// TIA Portal project "PLC_hackathon_2026_V21" (V21)

(* hardware
DEVICE "S71500/ET200MP station_1"  S7-1500 station
   slot 0: "Rail_0"  Rack  6ES7 590-1***0-0AA0
   slot 1: "PLC_1"  CPU 1515-2 PN  6ES7 515-2AM01-0AB0  V2.6
      slot 3: "CPU display_1"  6ES7591-1BA00-0AA0
DEVICE "PC-System_1"  SIMATIC PC station
   slot 0: "SIMATIC PC station"  Rail  SIMATIC PC-Station  V1.0
      slot 125: "Stationmanager"  Station_Manager  V6.0.4
   slot 1: "HMI_RT_1"  WinCC RT Advanced  6AV2 104-0xxxx-xxxx  17.0.0.0
      slot 33792: "Host interface"  Host interface
   slot 2: "IE general_1"  IE General  IE_CP  V8.2.0
*)

// ===== PLC "PLC_1"  CPU 1515-2 PN =====
// protected blocks, not shown: "Crane_manipulation"

VAR_GLOBAL   // PLC tag table "Default tag table"
   "x_position" AT %MB104 : SInt;
   "y_position" AT %MB105 : SInt;
   "bay_ID" AT %MB106 : USInt;
   "number_of_manipulations" AT %MD107 : UDInt;
   "time" AT %MD112 : Real;
END_VAR

VAR_GLOBAL   // PLC tag table "Crane_command"
   "new_x_position" AT %MB100 : SInt;   // X position for the move command
   "new_y_position" AT %MB101 : SInt;   // Y position for the move command
   "new_bay_ID" AT %MB102 : USInt;   // Bay ID for the move command
   "new_command_ID" AT %MB103 : USInt;   // ID of the command
END_VAR

TYPE "typeCmd"
   STRUCT
      Cmd : USInt;   // 0 none, 1 lift, 2 put down, 3 move to (X,Y,Bay), 10 reset
      X : SInt;   // 0..3 (for lift/put: current crane x)
      Y : SInt;   // 0..11 (for lift/put: current crane y)
      Bay : USInt;   // 0 ship, 1 yard
      Src : USInt;   // origin: 1 AUTO, 2 SEMI, 3 MANUAL, 4 INIT(reset)
      TrIdx : Int;   // plan transfer index (0 = not from plan)
      Phase : USInt;   // 0 move-to-src, 1 lift, 2 move-to-dst, 3 put (only if TrIdx>0)
   END_STRUCT;
END_TYPE

TYPE "typeTransfer"
   STRUCT
      Kind : USInt;   // 1 unload (Bay0->Bay1), 2 load (Bay1->Bay0)
      Id : UInt;   // container ID
      ListIdx : Int;   // index into UList (Kind 1) or LList (Kind 2)
      SrcX : SInt;
      SrcY : SInt;
      SrcBay : USInt;
      DstX : SInt;
      DstY : SInt;
      DstBay : USInt;
      CumT_ds : DInt;   // predicted total time after this transfer, deciseconds, incl. BaseT_ds
      CumM : DInt;   // predicted total manipulations after this transfer, incl. BaseM
   END_STRUCT;
END_TYPE

DATA_BLOCK "Current_state_of_Bay0"   // DB10
{ S7_Optimized_Access := 'TRUE' }
VERSION : 0.1
   VAR
      Bay0 : Array[0..3, 0..11] of UInt;
   END_VAR
BEGIN
   Bay0[0,0] := 123;
   Bay0[0,1] := 326;
   Bay0[0,2] := 987;
END_DATA_BLOCK

DATA_BLOCK "Current_state_of_Bay1"   // DB11
{ S7_Optimized_Access := 'TRUE' }
VERSION : 0.1
   VAR
      Bay1 : Array[0..3, 0..11] of UInt;
   END_VAR
BEGIN
   Bay1[0,1] := 246;
   Bay1[0,7] := 675;
   Bay1[1,5] := 777;
END_DATA_BLOCK

DATA_BLOCK "From_Bay0_to_Bay1"   // DB20
{ S7_Optimized_Access := 'TRUE' }
VERSION : 0.1
   VAR
      IDs_of_the_containers : Array[1..48] of UInt;
   END_VAR
BEGIN
   IDs_of_the_containers[12] := 0;
   IDs_of_the_containers[18] := 0;
   IDs_of_the_containers[4] := 444;
   IDs_of_the_containers[1] := 111;
   IDs_of_the_containers[2] := 222;
   IDs_of_the_containers[3] := 333;
   IDs_of_the_containers[5] := 555;
   IDs_of_the_containers[6] := 666;
   IDs_of_the_containers[7] := 777;
END_DATA_BLOCK

DATA_BLOCK "From_Bay1_to_Bay0"   // DB21
{ S7_Optimized_Access := 'TRUE' }
VERSION : 0.1
   VAR
      Bay1_IDs_of_the_containers : Array[1..48] of UInt;
   END_VAR
BEGIN
   Bay1_IDs_of_the_containers[15] := 0;
   Bay1_IDs_of_the_containers[22] := 0;
   Bay1_IDs_of_the_containers[1] := 123;
   Bay1_IDs_of_the_containers[2] := 124;
   Bay1_IDs_of_the_containers[3] := 125;
END_DATA_BLOCK

DATA_BLOCK "World"   // DB100
{ S7_Optimized_Access := 'TRUE' }
VERSION : 0.1
   VAR
      Bay0 : Array[0..3, 0..11] of UInt;   // working copy of the ship (FB10 INIT copy / OB30 lift-put effect)
      Bay1 : Array[0..3, 0..11] of UInt;   // working copy of the yard
      CraneX : SInt;   // crane x after last completed command
      CraneY : SInt;
      CraneBay : USInt := 1;
      Carried : UInt;   // ID on the hook (0 = none)
      Busy : Bool;   // command issued to FB1, not finished yet
      BusyTicks : Int;   // OB30 ticks since issue (watchdog)
      ActCmd : "typeCmd";   // command currently executing
      NextCmd : "typeCmd";   // staged command (valid when CmdReady)
      CmdReady : Bool;   // handshake: FB10 sets (last) / OB30 clears
      Permit : Bool;   // OB30 may issue NextCmd
      DoneSeq : UDInt;   // +1 per completed command
      LastDone : "typeCmd";   // last completed command
      Fault : Word;   // OB30-detected alarms (bit = alarm bit)
      FaultCmd : "typeCmd";   // command rejected by CheckCmd
      UList : Array[1..48] of UInt;   // copy of DB20 (unload list)
      UState : Array[1..48] of USInt;   // 0 pending, 1 done, 2 skipped
      LList : Array[1..48] of UInt;   // copy of DB21 (load list)
      LState : Array[1..48] of USInt;   // as UState
      N : Int;   // non-zero entries in DB20 + DB21 (for J)
      Plan : Array[1..96] of "typeTransfer";   // written by the planner
      PlanLen : Int;
      PlanValid : Bool;
      PlanVariant : Int;
      PredT_ds : DInt;
      PredM : DInt;
      PredJ : Real;
      BaseT_ds : DInt;   // ROUND(T*10) at plan request
      BaseM : DInt;   // M at plan request
      PlanIdx : Int := 1;   // done pointer: transfer being executed
      Phase : USInt;   // done pointer: next phase of PlanIdx to complete
      StageIdx : Int := 1;   // staging cursor (transfer)
      StagePhase : USInt;   // staging cursor (phase)
      BalL : Int;   // ship count x in {0,1}
      BalR : Int;   // ship count x in {2,3}
      BalF : Int;   // ship count y in 0..5
      BalA : Int;   // ship count y in 6..11
      CfgOrderMode : USInt := 1;   // 0 free, 1 per-list order, 2 strict (set by FB10 from HMI_IF before each plan)
      CfgBalLimit : Int := 5;
      CfgBalMode : USInt;   // 0 x-halves only, 1 also y-halves
      CfgMMode : USInt := 0;   // manipulation count model (CONTRACT 4.1); v1.7: 0 = spec rule (diagonal = 2), 2 = FB1 (+1 per move command)
      CfgVariants : Int := 4;
      CfgAlpha : Array[1..4] of Int;   // v1.7: retuned for CfgMMode 0 (v1.3 mode 2: [0, 100, 200, 300])
      CfgStepsPerCall : Int := 1;
      CfgTimeoutTicks : Int := 10;   // FB1 watchdog in OB30 ticks (1 s)
      OB30Ticks : UDInt;
      MSpec : UDInt;   // manipulations by the spec rule (OB30): +1 per changed axis, +1 lift/put ---- v1.3: improve phase (CONTRACT 4.8) and lower bound (4.9) ----
      CfgImproveEvals : DInt := 3000;   // local-search evaluations after the greedy (0 = off)
      CfgImproveDist : Int := 0;   // max |i-j| of a move (0 = unlimited)
      CfgImprovePerCall : Int := 1;   // evaluations per OB1 call (per-call work bound)
      PredJ0 : Real;   // J of the greedy winner before the improve phase
      LbT_ds : DInt;   // lower bound of the final T (incl. BaseT_ds), deciseconds
      LbM : DInt;   // lower bound of the final M (incl. BaseM)
      LbJ : Real;   // lower bound of J (no plan can be better)
      ImpEvals : DInt;   // improve phase: evaluations done (last plan)
      ImpAccepts : DInt;   // improve phase: accepted improvements (last plan) ---- v1.4: exact order feasibility (CONTRACT 4.10) and SLOT phase (4.11) ----
      CfgSlotSweeps : Int := 10;   // drop-cell local search sweeps after IMPROVE (0 = off)
      SlotAccepts : DInt;   // SLOT phase: accepted drop-cell changes (last plan)
      OrderFeasible : Bool;   // last plan job: the requested order mode is feasible (exact DP) ---- v1.5 (judge round 2 R2-J1): relaxed balance rule on a ship that starts out of balance ----
      BalCeil : Int;   // 0 = step rule; > CfgBalLimit: while |L-R| > CfgBalLimit a step may go up to BalCeil ---- v1.6 (judge round 3 R3-E3): relaxed ceiling search ----
      CfgRelaxMin : Bool;   // FALSE: relaxed fallback uses BalCeil = start imbalance at once; TRUE: ascending CfgBalLimit+1 .. start imbalance (smallest feasible, costs J)
   END_VAR
BEGIN
   CfgAlpha[1] := 0;
   CfgAlpha[2] := 75;
   CfgAlpha[3] := 125;
   CfgAlpha[4] := 200;
END_DATA_BLOCK

DATA_BLOCK "HMI_IF"   // DB101
{ S7_Optimized_Access := 'TRUE' }
VERSION : 0.1
// ---- Buttons / inputs (HMI writes; FB10 resets button bits after evaluating them) ----
   VAR
      SwOn : Bool;   // main switch level (HMI InvertBit), TRUE = ON
      BtnInit : Bool;   // INITIAL STATE (POCETNO STANJE)
      BtnAuto : Bool;
      BtnSemi : Bool;
      BtnManual : Bool;
      BtnStart : Bool;
      BtnStop : Bool;
      BtnAck : Bool;
      BtnStep : Bool;   // SEMI: run the next manipulation
      BtnManExec : Bool;   // MANUAL: execute ManCmd
      ManCmd : USInt;   // 1 lift, 2 put down, 3 move, 10 reset
      ManX : SInt;   // 0..3
      ManY : SInt;   // 0..11
      ManBay : USInt;   // 0 ship, 1 yard
      CfgOrderMode : USInt := 1;   // 0 free, 1 per-list order (default, hedge), 2 strict; FB10 falls back 2->1->0 if infeasible
      CfgSemiPerTransfer : Bool;   // SEMI click = one command (FALSE) or one transfer (TRUE)
      CfgBalMode : USInt;   // 0 x-halves, 1 also y-halves
      AlarmHmiAck : Word;   // WinCC 'Acknowledgement tag': alarm acknowledged in the alarm view (= POTVRDA); FB10 resets it ---- Indicators (FB10 writes every OB1 cycle) ----
      State : USInt;   // 0 OFF,1 INIT,2 READY,3 RUNNING,4 PAUSED,5 ALARM,6 DONE,7 PLANNING
      Mode : USInt := 1;   // 1 AUTO, 2 SEMI, 3 MANUAL
      LampOn : Bool;
      LampOff : Bool;
      LampReady : Bool;
      LampAuto : Bool;
      LampSemi : Bool;
      LampManual : Bool;
      LampRunning : Bool;
      LampAlarm : Bool;
      LampDone : Bool;
      Initialized : Bool;
      CraneBusy : Bool;
      Planning : Bool;
      StepWaiting : Bool;   // SEMI is waiting for a click
      "M" : UDInt;   // v1.7: M by the spec rule (x and y change = 2) = World.MSpec (primary)
      T : Real;   // = "time" (MD112) working time [s]
      J : Real;   // v1.7: 0.5*T/(76*N) + 0.5*M/(4*N) with the spec M (primary)
      MSpec : UDInt;   // = M (spec rule, computed in OB30); kept for compatibility
      JSpec : Real;   // = J (spec rule); kept for compatibility
      MFb1 : UDInt;   // v1.7: FB1's own counter "number_of_manipulations" (MD107, +1 per command)
      JFb1 : Real;   // v1.7: J with MFb1 (secondary)
      OrderModeAct : USInt;   // order mode actually used by the last plan (after fallback)
      OrderFallback : Bool;   // v1.4: preferred order/balance mode infeasible, plan uses a weaker one
      SlotAccepts : DInt;   // v1.4: SLOT phase accepted drop-cell changes (last plan)
      N : Int;
      PredM : DInt;
      PredT : Real;
      PredJ : Real;
      PredJ0 : Real;   // v1.3: greedy J before the improve phase
      LbJ : Real;   // v1.3: lower bound of J (no plan can be better)
      GapPct : Real;   // v1.3: (PredJ / LbJ - 1) * 100
      ImpGainPct : Real;   // v1.3: (1 - PredJ / PredJ0) * 100 = gain of the improve phase
      ImpEvals : DInt;   // v1.3: improve-phase evaluations of the last plan
      PlanProgress : Int;   // v1.3: planner progress 0..100 % (improve phase)
      PlanVariant : Int;
      TrDone : Int;
      TrTotal : Int;
      UDone : Int;
      UTotal : Int;
      LDone : Int;
      LTotal : Int;
      CraneX : SInt;
      CraneY : SInt;
      CraneBay : USInt;
      CraneGX : Int;   // global column: x+6 if bay 0 else x (0..9)
      Carried : UInt;
      CurCmd : USInt;
      CurX : SInt;
      CurY : SInt;
      CurBay : USInt;
      CurId : UInt;
      CurKind : USInt;   // 1 unload, 2 load, 0 none
      CurPhase : USInt;
      Cell0 : Array[0..47] of UInt;   // Bay0 IDs, index x*12+y
      Cell1 : Array[0..47] of UInt;   // Bay1 IDs, index x*12+y
      CellSt0 : Array[0..47] of USInt;   // colour code 0..7
      CellSt1 : Array[0..47] of USInt;
      UList : Array[1..48] of UInt;
      LList : Array[1..48] of UInt;
      UState : Array[1..48] of USInt;   // 0 pending, 1 done, 2 skipped, 3 in progress
      LState : Array[1..48] of USInt;
      BalL : Int;
      BalR : Int;
      BalDiff : Int;   // BalL - BalR
      BalF : Int;
      BalA : Int;
      BalOk : Bool;   // |BalDiff| <= 5
      AlarmWord : Word;   // alarm bits (CONTRACT 3.3)
      AlarmAckWord : Word;   // WinCC 'PLC acknowledgement tag' = NOT AlarmWord (one ACK clears PLC and HMI)
      AlarmId : UInt;
      AlarmWord2 : Word;   // v1.4: extra alarm bits: bit 0 = list order abandoned (warning); v1.5 bit 1 = relaxed balance rule (ship loaded unbalanced)
      AlarmUId : UInt;   // v1.4: first unload-list ID that is not in Bay 0 (alarm bit 3)
      AlarmUCnt : Int;   // number of such IDs
      AlarmLId : UInt;   // v1.4: first load-list ID that is not in Bay 1 (alarm bit 4)
      AlarmLCnt : Int;
      AlarmX : SInt;
      AlarmY : SInt;
      AlarmBay : USInt;
      AlarmHist : Array[0..15] of Int;   // alarm bit numbers of the last 16 raises, [0] newest
      AlarmHistSeq : UDInt;
      OB30Ticks : UDInt;
      Heartbeat : Bool;   // toggles each OB30 tick
   END_VAR
BEGIN
END_DATA_BLOCK

DATA_BLOCK "Crane_Control_DB"   // DB110
{ S7_Optimized_Access := 'TRUE' }
VERSION : 0.1
// stored: InstanceOfName Crane_Control
"Crane_Control"
BEGIN
END_DATA_BLOCK

// folder: Constants

DATA_BLOCK "Global_constants"   // DB1
{ S7_Optimized_Access := 'TRUE' }
VERSION : 0.1
   VAR
      container_width_in_m : Real := 2.3;   // Container width in meters
      container_length_in_m : Real := 6.0;   // Container length in meters
      velocity_of_the_crane_in_m_per_s : Real := 1.0;   // Velocity of the crane in meters per second
      time_to_lift_a_container_in_s : Real := 20.0;   // Time needed to lower the hook, hook up a container and lift it in seconds
      time_to_put_down_a_container_in_s : Real := 20.0;   // Time needed to put down a container, release it, and lift up the hook in seconds
   END_VAR
BEGIN
END_DATA_BLOCK

// folder: (top level)

FUNCTION_BLOCK "Crane_Control"   // FB10, SCL
TITLE = Container crane control (FB10, called from OB1)
{ S7_Optimized_Access := 'TRUE' }
VERSION : 0.1
// FB10 decides WHAT the crane does; OB30 decides WHEN (CONTRACT 3.4).
//   - HMI buttons, modes AUTO / SEMI-AUTO / MANUAL
//   - state machine OFF / INIT / READY / RUNNING / PAUSED / ALARM / DONE / PLANNING
//   - INIT: reset FB1, copy DB10/DB11, validate lists and IDs, call the planner
//   - stages plan commands into "World".NextCmd (handshake CmdReady / Permit)
//   - tracks progress (done pointer), list states, ship balance, alarms
//   - writes every indicator of "HMI_IF"
//   FB10 never calls FB1 and never writes MB100..MB103; FB1 tags are read-only here.
   VAR
      Planner : "Crane_Planner";   // planning algorithm (FB11, CONTRACT 4)
      PlanReq : Bool;   // Req input of the planner
      PlanFinished : Bool;   // planner job ended, result not yet consumed
      PlanOk : Bool;
      PlanErr : Int;
      PlanStep : Int;   // PLANNING sub-step
      PlanCrX : SInt;   // crane position at plan request
      PlanCrY : SInt;
      PlanCrBay : USInt;
      FirstPh : Array[1..96] of USInt;   // first phase of each transfer (1 = move-to-src skipped)
      State : USInt;   // 0 OFF,1 INIT,2 READY,3 RUNNING,4 PAUSED,5 ALARM,6 DONE,7 PLANNING
      PrevState : USInt;   // state to return to after ALARM + ACK
      OffState : USInt;   // state before OFF
      Mode : USInt := 1;   // 1 AUTO, 2 SEMI, 3 MANUAL
      PendMode : USInt;   // mode press waiting to be applied
      Initialized : Bool;
      InitStep : Int;   // INIT sub-step
      InitSeq : UDInt;   // DoneSeq when the INIT reset was staged
      SeenSeq : UDInt;   // last "World".DoneSeq processed
      Resync : Bool;   // re-align staging cursor to done pointer before staging
      SemiTokens : Int;   // SEMI: commands still allowed by BtnStep
      AlarmLatch : Word;   // latched alarm bits (CONTRACT 3.3)
      AlarmPrev : Word;   // for raise-edge detection (history)
      AlarmHistM : Array[0..15] of UDInt;   // M at each history entry (parallel to HMI_IF.AlarmHist)
      AlarmHistT : Array[0..15] of Real;   // T [s] at each history entry
      FirstScan : Bool := TRUE;
      Snap0 : Array[0..3, 0..11] of UInt;   // DB10 as last seen: external online edits are adopted into World
      Snap1 : Array[0..3, 0..11] of UInt;   // DB11 as last seen
      PendStep : Bool;   // SEMI: latched NEXT STEP click (kept while FB1 is busy)
      ReplanAfterPut : Bool;   // destination re-targeted after ACK: replan after that put
      CfgOrdHmi : USInt := 1;   // CfgOrderMode last taken from the HMI (preferred mode)
      CfgBalHmi : USInt;   // CfgBalMode last taken from the HMI
      OrdFallback : Bool;   // next plan request is a fallback retry (keep World.Cfg*) v1.4: DB10/DB11 are kept as the live state; copy of the loaded data for POÄŒETNO STANJE
      InitBay0 : Array[0..3, 0..11] of UInt;
      InitBay1 : Array[0..3, 0..11] of UInt;
      HaveInit : Bool;   // InitBay0/1 valid
      ExtEdit : Bool;   // v1.6: not used any more (NewCnt / ObstCnt), kept for the interface
      NoCellWarn : Bool;   // v1.5: bit 7 raised by the ACK re-target (MANUAL needed): not blocking
      BalD0 : Int;   // v1.5 (R2-J1): |L-R| of the ship as loaded at INIT v1.6 (judge round 3 R3-E1 / R3-J1): obstacle edits during a job are not a new data set
      JobActive : Bool;   // a plan or MANUAL command completed since the last INIT
      EditMark : Array[0..95] of Bool;   // cell (bay*48 + x*12 + y) edited online since the last INIT
      EditNew : Array[0..95] of Bool;   // ... and that edit was made while no job was in progress
      EditVal : Array[0..95] of UInt;   // value of the cell before the edit (written back = unmarked)
      NewCnt : Int;   // marked cells edited with no job in progress (new data)
      ObstCnt : Int;   // marked cells edited during a job (obstacles)
   END_VAR
   VAR_TEMP
      visSt0 : Array[0..47] of USInt;   // display colours built privately
      visSt1 : Array[0..47] of USInt;
      bInit : Bool;   // button snapshots (HMI bits are reset at once)
      bAuto : Bool;
      bSemi : Bool;
      bManual : Bool;
      bStart : Bool;
      bStop : Bool;
      bAck : Bool;
      bStep : Bool;
      bManExec : Bool;
      i : Int;
      j : Int;
      k : Int;
      x : Int;
      y : Int;
      "b" : Int;
      id : UInt;
      found : Bool;
      found0 : Bool;
      found1 : Bool;
      cnt : Int;
      cnt2 : Int;
      pu : Int;
      pl : Int;
      seq : UDInt;
      last : "typeCmd";
      cur : "typeCmd";
      blocking : Bool;
      hadFault : Bool;
      carriedOk : Bool;
      newBits : Word;
      newFault : Word;
      tc : Array[0..95] of UInt;   // INIT: all cells, index bay*48 + x*12 + y
      tl : Array[1..96] of UInt;   // INIT: UList (1..48) then LList (49..96)
      ts : Array[1..96] of USInt;   // INIT: states of tl
      rN : Real;
      curValid : Bool;
      tr : "typeTransfer";
      unbal : Bool;   // ship out of balance now (alarm bit 0 condition)
      semiGo : Bool;   // SEMI NEXT STEP in READY / PAUSED = START + one step
      faultWas : Word;   // World.Fault at ACK
      planPut : Bool;   // completed PUT belongs to the plan
      bestT : Int;   // re-target: best travel time [ds]
      bestX : Int;
      bestY : Int;
      candT : Int;
      nL : Int;
      nR : Int;
      nF : Int;
      nA : Int;
      okBal : Bool;
      dstB : USInt;
      noCell : Bool;   // ACK: rejected plan put could not be re-targeted
      extE : Bool;   // INIT: DB10/DB11 differ from the last mirrored state
      noJob : Bool;   // v1.6: no job in progress (an online edit is new data)
      dbv : UInt;   // v1.6 region 2a: DB10/DB11 cell
      snv : UInt;   // Snap cell
      wv : UInt;   // World cell v1.6 (judge round 3 R3-E2): order feasibility of the ACK re-target (bit-parallel FtMask[0,0])
      ft0 : DWord;   // bit L: the remaining lists stay feasible from L ship containers in x 0..1
      ftNu : Int;   // remaining pending unloads (list order)
      ftNl : Int;   // remaining pending loads (without the one on the hook)
      ftS0 : Int;   // ship count after the put
      ftY0 : Int;   // yard count
      ftCeil : Int;   // ceiling of this try: 0 step rule, > 0 relaxed, -1 skip, -2 no filter
      ftTry : Int;
      ftUse : Bool;   // filter possible (ship put, preferred order 1 / 2)
      ftSide : Array[1..48] of Bool;   // pending unload i (list order) stands in x 0..1
      ftPrev : Array[0..48] of DWord;   // FtMask row i + 1
      ftCur : Array[0..48] of DWord;   // FtMask row i
      ftK : Array[0..4, 0..48] of DWord;   // per ship total: 0 end state, 1 unload left, 2 unload right, 3 load left, 4 load right
      ftTot : Int;
      ftL : Int;
      ftR : Int;
      ftD : Int;
      ftD2 : Int;
      ftM : DWord;
      ftBit : DWord;
      listsNew : Bool;   // v1.6 INIT: DB20/DB21 differ from the lists of the last load
   END_VAR
BEGIN
   REGION 0 First scan after PLC start
       IF #FirstScan THEN
           FOR #i := 0 TO 15 DO
               "HMI_IF".AlarmHist[#i] := -1;      // -1 = empty history entry
           END_FOR;
           #Mode := 1;                            // default AUTO
           #State := 0;
           #FirstScan := FALSE;
       END_IF;
   END_REGION

   REGION 1 HMI buttons: snapshot and reset
       #bInit := "HMI_IF".BtnInit;       "HMI_IF".BtnInit := FALSE;
       #bAuto := "HMI_IF".BtnAuto;       "HMI_IF".BtnAuto := FALSE;
       #bSemi := "HMI_IF".BtnSemi;       "HMI_IF".BtnSemi := FALSE;
       #bManual := "HMI_IF".BtnManual;   "HMI_IF".BtnManual := FALSE;
       #bStart := "HMI_IF".BtnStart;     "HMI_IF".BtnStart := FALSE;
       #bStop := "HMI_IF".BtnStop;       "HMI_IF".BtnStop := FALSE;
       #bAck := "HMI_IF".BtnAck;         "HMI_IF".BtnAck := FALSE;
       #bStep := "HMI_IF".BtnStep;       "HMI_IF".BtnStep := FALSE;
       #bManExec := "HMI_IF".BtnManExec; "HMI_IF".BtnManExec := FALSE;
       // Alarm acknowledged in the WinCC alarm view ("Acknowledgement tag") = POTVRDA
       IF "HMI_IF".AlarmHmiAck <> 0 THEN
           #bAck := TRUE;
           "HMI_IF".AlarmHmiAck := 0;
       END_IF;
       // SEMI: a NEXT STEP click is latched until it can be executed (FB1 busy, planning, ...)
       IF #bStep AND #Mode = 2 THEN
           #PendStep := TRUE;
       END_IF;
   END_REGION

   REGION 2a DB10 / DB11 = live state: mirror our moves, adopt external online edits
       // After INIT our container model is World.Bay0/Bay1 (OB30 updates it after every lift / put).
       // Snap0/Snap1 = DB10/DB11 as last written or seen by this block.
       //  - DB10/DB11 cell <> Snap: changed online (watch table, HMI) -> taken over into World, so the
       //    OB30 pre-check "pick location empty / drop location occupied" acts on it and the grid shows it.
       //    v1.5: in every state such an edit counts as new input data for the next POÄŒETNO STANJE
       //    (ExtEdit, see INIT; judge round 2 R2-E2 / R2-J3). v1.6: see below.
       //  - else World cell <> Snap: the crane moved a container -> written into DB10/DB11, so the given
       //    "Current_state_of_Bay0/1" blocks always show the current yard (v1.4, judge round 1 R1-E2).
       //  v1.6 (judge round 3 R3-E1 / R3-J1): every edited cell is marked (EditMark, value before the edit in
       //  EditVal). An edit made while NO job is in progress (nothing executed since INIT, or DONE) is new
       //  data (NewCnt); an edit during a job (an obstacle written to provoke "drop location occupied") is
       //  an obstacle (ObstCnt). Writing the cell back to its value before the edit removes the mark again.
       //  INIT takes DB10/DB11 as the new yard only if NewCnt > 0, or the lists changed and ObstCnt > 0, or
       //  ObstCnt >= 8 (a whole data set typed in while paused); otherwise it restores the loaded yard.
       #extE := FALSE;
       #noJob := NOT #JobActive OR #State = 6 OR (#State = 5 AND #PrevState = 6) OR (#State = 0 AND #OffState = 6);
       IF #Initialized AND #State <> 1 THEN
           FOR #b := 0 TO 1 DO
               FOR #x := 0 TO 3 DO
                   FOR #y := 0 TO 11 DO
                       IF #b = 0 THEN
                           #dbv := "Current_state_of_Bay0".Bay0[#x, #y];
                           #snv := #Snap0[#x, #y];
                           #wv := "World".Bay0[#x, #y];
                       ELSE
                           #dbv := "Current_state_of_Bay1".Bay1[#x, #y];
                           #snv := #Snap1[#x, #y];
                           #wv := "World".Bay1[#x, #y];
                       END_IF;
                       #k := #b * 48 + #x * 12 + #y;
                       IF #dbv <> #snv THEN
                           // changed online -> adopt into World, mark the cell
                           IF NOT #EditMark[#k] THEN
                               #EditMark[#k] := TRUE;
                               #EditVal[#k] := #snv;
                               #EditNew[#k] := #noJob;
                               IF #noJob THEN
                                   #NewCnt := #NewCnt + 1;
                               ELSE
                                   #ObstCnt := #ObstCnt + 1;
                               END_IF;
                           ELSIF #dbv = #EditVal[#k] THEN
                               #EditMark[#k] := FALSE;    // written back: no longer an edit
                               IF #EditNew[#k] THEN
                                   #NewCnt := #NewCnt - 1;
                               ELSE
                                   #ObstCnt := #ObstCnt - 1;
                               END_IF;
                           END_IF;
                           #extE := TRUE;
                           IF #b = 0 THEN
                               #Snap0[#x, #y] := #dbv;
                               "World".Bay0[#x, #y] := #dbv;
                           ELSE
                               #Snap1[#x, #y] := #dbv;
                               "World".Bay1[#x, #y] := #dbv;
                           END_IF;
                       ELSIF #wv <> #snv THEN
                           // the crane moved a container -> mirror it into DB10/DB11
                           IF #b = 0 THEN
                               #Snap0[#x, #y] := #wv;
                               "Current_state_of_Bay0".Bay0[#x, #y] := #wv;
                           ELSE
                               #Snap1[#x, #y] := #wv;
                               "Current_state_of_Bay1".Bay1[#x, #y] := #wv;
                           END_IF;
                       END_IF;
                   END_FOR;
               END_FOR;
           END_FOR;
           // v1.5 (judge round 2 R2-E2): an adopted edit while not running invalidates the plan, so the
           // next START replans on the edited yard instead of running a stale plan (with an empty hook;
           // with a load the plan is kept so the transfer in progress can be finished).
           IF #extE AND (#State = 0 OR #State = 2 OR #State = 4 OR #State = 5 OR #State = 6)
               AND "World".Carried = 0
           THEN
               "World".PlanValid := FALSE;
           END_IF;
       END_IF;
   END_REGION

   REGION 2 Planner call (multi-instance; runs a few greedy steps per OB1 cycle)
       #Planner(Req := #PlanReq);
       IF #PlanReq AND (#Planner.Done OR #Planner.Error) THEN
           #PlanFinished := TRUE;
           #PlanOk := #Planner.Done AND NOT #Planner.Error;
           #PlanErr := #Planner.ErrCode;
           #PlanReq := FALSE;                     // falling edge clears Done/Error
       END_IF;
   END_REGION

   REGION 3 Completed commands: done pointer, list states, manual commands
       // Read DoneSeq, then LastDone, then DoneSeq again: if OB30 ran in between,
       // skip this cycle and take a consistent snapshot in the next one.
       #seq := "World".DoneSeq;
       #last := "World".LastDone;
       IF #seq <> #SeenSeq AND #seq = "World".DoneSeq THEN
           #SeenSeq := #seq;
           IF #last.Src >= 1 AND #last.Src <= 3 THEN
               #JobActive := TRUE;                // v1.6: from now on online edits are obstacles
           END_IF;

           // Plan command finished: advance the done pointer (PlanIdx / Phase)
           IF (#last.Src = 1 OR #last.Src = 2) AND "World".PlanValid
               AND #last.TrIdx = "World".PlanIdx AND #last.Phase = "World".Phase
           THEN
               IF "World".Phase >= 3 THEN
                   "World".PlanIdx := "World".PlanIdx + 1;
                   IF "World".PlanIdx >= 1 AND "World".PlanIdx <= "World".PlanLen AND "World".PlanIdx <= 96 THEN
                       "World".Phase := #FirstPh["World".PlanIdx];
                   ELSE
                       "World".Phase := 0;
                   END_IF;
               ELSE
                   "World".Phase := "World".Phase + 1;
               END_IF;
           END_IF;

           // Manual command finished: the plan no longer matches the yard -> replan on START
           IF #last.Src = 3 THEN
               "World".PlanValid := FALSE;
               IF #State = 6 THEN
                   #State := 4;                   // DONE -> PAUSED (lists may be pending again)
               END_IF;
               IF #State <> 3 THEN
                   "World".Permit := FALSE;
               END_IF;
           END_IF;

           // After every PUT: update the list states
           IF #last.Cmd = 2 THEN
               // Plan put (AUTO / SEMI): exactly its own list entry is done (robust against
               // duplicate IDs, which INIT accepts with a bit 6 warning)
               #planPut := FALSE;
               IF (#last.Src = 1 OR #last.Src = 2) AND #last.Phase = 3 AND #last.TrIdx >= 1 AND #last.TrIdx <= 96
                   AND #last.X >= 0 AND #last.X <= 3 AND #last.Y >= 0 AND #last.Y <= 11 AND #last.Bay <= 1
               THEN
                   #tr := "World".Plan[#last.TrIdx];
                   IF #last.Bay = 0 THEN
                       #id := "World".Bay0[SINT_TO_INT(#last.X), SINT_TO_INT(#last.Y)];
                   ELSE
                       #id := "World".Bay1[SINT_TO_INT(#last.X), SINT_TO_INT(#last.Y)];
                   END_IF;
                   IF #id <> 0 AND #id = #tr.Id AND #last.Bay = #tr.DstBay AND #tr.ListIdx >= 1 AND #tr.ListIdx <= 48 THEN
                       IF #tr.Kind = 1 AND "World".UState[#tr.ListIdx] = 0 THEN
                           "World".UState[#tr.ListIdx] := 1;
                           #planPut := TRUE;
                       ELSIF #tr.Kind = 2 AND "World".LState[#tr.ListIdx] = 0 THEN
                           "World".LState[#tr.ListIdx] := 1;
                           #planPut := TRUE;
                       END_IF;
                   END_IF;
                   // the destination was re-targeted after a "drop occupied" ACK: replan now
                   IF #ReplanAfterPut THEN
                       #ReplanAfterPut := FALSE;
                       "World".PlanValid := FALSE;
                   END_IF;
               END_IF;

               // MANUAL put: presence check. Done only if the ID is in the destination bay and no
               // longer in the source bay; pending again only in the opposite case (an ID that is in
               // both bays, i.e. a duplicate, never changes the state).
               IF NOT #planPut THEN
                   FOR #i := 1 TO 48 DO
                       #id := "World".UList[#i];
                       IF #id <> 0 AND "World".UState[#i] <= 1 THEN
                           #found0 := FALSE;
                           #found1 := FALSE;
                           FOR #x := 0 TO 3 DO
                               FOR #y := 0 TO 11 DO
                                   IF "World".Bay0[#x, #y] = #id THEN #found0 := TRUE; END_IF;
                                   IF "World".Bay1[#x, #y] = #id THEN #found1 := TRUE; END_IF;
                               END_FOR;
                           END_FOR;
                           IF "World".UState[#i] = 0 AND #found1 AND NOT #found0 THEN
                               "World".UState[#i] := 1;
                           ELSIF "World".UState[#i] = 1 AND #found0 AND NOT #found1 THEN
                               "World".UState[#i] := 0;
                           END_IF;
                       END_IF;
                       #id := "World".LList[#i];
                       IF #id <> 0 AND "World".LState[#i] <= 1 THEN
                           #found0 := FALSE;
                           #found1 := FALSE;
                           FOR #x := 0 TO 3 DO
                               FOR #y := 0 TO 11 DO
                                   IF "World".Bay0[#x, #y] = #id THEN #found0 := TRUE; END_IF;
                                   IF "World".Bay1[#x, #y] = #id THEN #found1 := TRUE; END_IF;
                               END_FOR;
                           END_FOR;
                           IF "World".LState[#i] = 0 AND #found0 AND NOT #found1 THEN
                               "World".LState[#i] := 1;
                           ELSIF "World".LState[#i] = 1 AND #found1 AND NOT #found0 THEN
                               "World".LState[#i] := 0;
                           END_IF;
                       END_IF;
                   END_FOR;
               END_IF;
           END_IF;
       END_IF;
   END_REGION

   REGION 4 Ship balance (continuous) and configuration
       "World".BalL := 0;
       "World".BalR := 0;
       "World".BalF := 0;
       "World".BalA := 0;
       FOR #x := 0 TO 3 DO
           FOR #y := 0 TO 11 DO
               IF "World".Bay0[#x, #y] <> 0 THEN
                   IF #x <= 1 THEN
                       "World".BalL := "World".BalL + 1;
                   ELSE
                       "World".BalR := "World".BalR + 1;
                   END_IF;
                   IF #y <= 5 THEN
                       "World".BalF := "World".BalF + 1;
                   ELSE
                       "World".BalA := "World".BalA + 1;
                   END_IF;
               END_IF;
           END_FOR;
       END_FOR;
       // Alarm bit 0 while the ship is out of balance (warning; CheckCmd in OB30
       // blocks every lift/put that would make it worse)
       #unbal := #Initialized AND (ABS("World".BalL - "World".BalR) > "World".CfgBalLimit
           OR ("World".CfgBalMode = 1 AND ABS("World".BalF - "World".BalA) > "World".CfgBalLimit));
       IF #unbal THEN
           #AlarmLatch := #AlarmLatch OR WORD#16#0001;
       END_IF;

       // Planner configuration from the HMI: only while nothing runs and the hook is empty
       // (a change takes effect at the next transfer boundary; a replan needs an empty hook).
       // CfgOrdHmi / CfgBalHmi are the preferred modes; World.Cfg* may be lowered by the
       // infeasibility fallback and are set back to the preferred modes before every plan request.
       IF #State <> 1 AND #State <> 3 AND #State <> 7 AND "World".Carried = 0 AND NOT "World".Busy THEN
           IF "HMI_IF".CfgOrderMode <= 2 AND "HMI_IF".CfgOrderMode <> #CfgOrdHmi THEN
               #CfgOrdHmi := "HMI_IF".CfgOrderMode;
               "World".CfgOrderMode := #CfgOrdHmi;
               "World".PlanValid := FALSE;
           END_IF;
           IF "HMI_IF".CfgBalMode <= 1 AND "HMI_IF".CfgBalMode <> #CfgBalHmi THEN
               #CfgBalHmi := "HMI_IF".CfgBalMode;
               "World".CfgBalMode := #CfgBalHmi;
               "World".PlanValid := FALSE;
           END_IF;
       END_IF;
   END_REGION

   REGION 5 Alarms raised by OB30 (World.Fault) and ACK
       // New OB30 faults: take over and remember where they happened
       #newFault := "World".Fault AND NOT #AlarmLatch;
       IF #newFault <> 0 THEN
           IF (#newFault AND WORD#16#4400) <> 0 THEN      // bit 10 timeout / bit 14 position
               #cur := "World".ActCmd;
           ELSE
               #cur := "World".FaultCmd;
           END_IF;
           "HMI_IF".AlarmX := #cur.X;
           "HMI_IF".AlarmY := #cur.Y;
           "HMI_IF".AlarmBay := #cur.Bay;
           "HMI_IF".AlarmId := "World".Carried;
           IF "World".Carried = 0 AND #cur.X >= 0 AND #cur.X <= 3 AND #cur.Y >= 0 AND #cur.Y <= 11 THEN
               IF #cur.Bay = 0 THEN
                   "HMI_IF".AlarmId := "World".Bay0[SINT_TO_INT(#cur.X), SINT_TO_INT(#cur.Y)];
               ELSIF #cur.Bay = 1 THEN
                   "HMI_IF".AlarmId := "World".Bay1[SINT_TO_INT(#cur.X), SINT_TO_INT(#cur.Y)];
               END_IF;
           END_IF;
       END_IF;
       #AlarmLatch := #AlarmLatch OR "World".Fault;

       // ACK: clear all latched bits; bits whose cause persists are raised again.
       // An ACK in the same cycle as a new OB30 fault is ignored: the fault must first stop the
       // system (ALARM) and enter the history; the operator acknowledges it afterwards.
       // The imbalance bit 0 stays latched while the ship is still out of balance (no new history entry).
       IF #bAck AND #newFault = 0 THEN
           #NoCellWarn := FALSE;
           #faultWas := "World".Fault;
           #hadFault := #faultWas <> 0;
           "World".Fault := "World".Fault AND NOT #faultWas;
           IF #unbal THEN
               #AlarmLatch := WORD#16#0001;
           ELSE
               #AlarmLatch := 0;
           END_IF;
           "HMI_IF".AlarmId := 0;

           // "Drop location occupied" (bit 2) or "put would unbalance the ship" (bit 0, CheckCmd 100)
           // for a plan put with the container on the hook: put it on the nearest free cell of the same
           // bay that keeps the ship balanced, then replan ("nakon potvrde sustav nastavlja s radom").
           // v1.4: bit 0 added; with no such cell the system PAUSES (bit 7, MANUAL needed) instead of
           // re-staging the same rejected put (endless ALARM / ACK loop, judge round 1 R1-E3).
           #noCell := FALSE;
           IF (#faultWas AND WORD#16#0005) <> 0 AND "World".Carried <> 0 AND "World".PlanValid
               AND "World".FaultCmd.Cmd = 2 AND ("World".FaultCmd.Src = 1 OR "World".FaultCmd.Src = 2)
               AND "World".PlanIdx >= 1 AND "World".PlanIdx <= "World".PlanLen AND "World".PlanIdx <= 96
               AND "World".Phase = 3 AND "World".CraneBay <= 1
           THEN
               #dstB := "World".CraneBay;
               // v1.6 (judge round 3 R3-E2): for a SHIP put, prefer the cells whose side keeps the remaining
               // lists feasible in the preferred order (exact FtMask[0,0] of the state after the put, the same
               // table as FB11, here bit-parallel: try 1 step rule, try 2 relaxed ceiling BalD0). Try 3 = the
               // v1.4 rule (nearest balance-safe cell) when no cell keeps the order. Python reference:
               // tools/fb10_init_model.retarget() / ft00().
               #ftUse := #dstB = 0 AND #CfgOrdHmi > 0;
               #ftNu := 0;
               #ftNl := 0;
               #ftS0 := "World".BalL + "World".BalR + 1;
               #ftY0 := 0;
               IF #ftUse THEN
                   FOR #x := 0 TO 3 DO
                       FOR #y := 0 TO 11 DO
                           IF "World".Bay1[#x, #y] <> 0 THEN
                               #ftY0 := #ftY0 + 1;
                           END_IF;
                       END_FOR;
                   END_FOR;
                   FOR #i := 1 TO 48 DO
                       #id := "World".UList[#i];
                       IF #id <> 0 AND "World".UState[#i] = 0 THEN
                           #found := FALSE;
                           FOR #x := 0 TO 3 DO
                               FOR #y := 0 TO 11 DO
                                   IF NOT #found AND "World".Bay0[#x, #y] = #id THEN
                                       #found := TRUE;
                                       #ftNu := #ftNu + 1;
                                       #ftSide[#ftNu] := #x <= 1;
                                   END_IF;
                               END_FOR;
                           END_FOR;
                       END_IF;
                       #id := "World".LList[#i];
                       IF #id <> 0 AND "World".LState[#i] = 0
                           AND NOT ("World".Plan["World".PlanIdx].Kind = 2 AND "World".Plan["World".PlanIdx].ListIdx = #i)
                       THEN
                           #found := FALSE;
                           FOR #x := 0 TO 3 DO
                               FOR #y := 0 TO 11 DO
                                   IF "World".Bay1[#x, #y] = #id THEN
                                       #found := TRUE;
                                   END_IF;
                               END_FOR;
                           END_FOR;
                           IF #found THEN
                               #ftNl := #ftNl + 1;
                           END_IF;
                       END_IF;
                   END_FOR;
               END_IF;
               #bestX := -1;
               #bestY := -1;
               FOR #ftTry := 1 TO 3 DO
                   IF #bestX < 0 THEN
                       #ftCeil := -1;
                       IF #ftTry = 1 AND #ftUse THEN
                           #ftCeil := 0;
                       ELSIF #ftTry = 2 AND #ftUse AND #BalD0 > "World".CfgBalLimit THEN
                           #ftCeil := #BalD0;
                       ELSIF #ftTry = 3 THEN
                           #ftCeil := -2;
                       END_IF;
                       IF #ftCeil >= 0 THEN
                           // move masks per ship total (bit L, R = tot - L)
                           FOR #ftTot := 0 TO 48 DO
                               FOR #k := 0 TO 4 DO
                                   #ftK[#k, #ftTot] := DWORD#16#0;
                               END_FOR;
                               FOR #ftL := 0 TO 24 DO
                                   #ftR := #ftTot - #ftL;
                                   IF #ftR >= 0 AND #ftR <= 24 THEN
                                       #ftBit := SHL(IN := DWORD#16#1, N := INT_TO_USINT(#ftL));
                                       #ftD := ABS(#ftL - #ftR);
                                       IF #ftCeil = 0 OR #ftD <= "World".CfgBalLimit THEN
                                           #ftK[0, #ftTot] := #ftK[0, #ftTot] OR #ftBit;     // end state (relaxed: balanced)
                                       END_IF;
                                       FOR #k := 1 TO 4 DO
                                           IF (#k = 1 AND #ftL >= 1) OR (#k = 2 AND #ftR >= 1)
                                               OR (#k = 3 AND #ftL <= 23) OR (#k = 4 AND #ftR <= 23)
                                           THEN
                                               IF #k = 1 THEN
                                                   #ftD2 := ABS(#ftL - 1 - #ftR);
                                               ELSIF #k = 2 THEN
                                                   #ftD2 := ABS(#ftL - #ftR + 1);
                                               ELSIF #k = 3 THEN
                                                   #ftD2 := ABS(#ftL + 1 - #ftR);
                                               ELSE
                                                   #ftD2 := ABS(#ftL - #ftR - 1);
                                               END_IF;
                                               IF #ftD2 <= "World".CfgBalLimit OR #ftD2 <= #ftD
                                                   OR (#ftD > "World".CfgBalLimit AND #ftD2 <= #ftCeil)
                                               THEN
                                                   #ftK[#k, #ftTot] := #ftK[#k, #ftTot] OR #ftBit;
                                               END_IF;
                                           END_IF;
                                       END_FOR;
                                   END_IF;
                               END_FOR;
                           END_FOR;
                           // FtMask rows i = ftNu .. 0 (two row buffers)
                           FOR #j := 0 TO 48 DO
                               #ftPrev[#j] := DWORD#16#0;
                               #ftCur[#j] := DWORD#16#0;
                           END_FOR;
                           FOR #i := #ftNu TO 0 BY -1 DO
                               FOR #j := #ftNl TO 0 BY -1 DO
                                   #ftTot := #ftS0 - #i + #j;
                                   #ftM := DWORD#16#0;
                                   IF #ftTot >= 0 AND #ftTot <= 48 THEN
                                       IF #i = #ftNu AND #j = #ftNl THEN
                                           #ftM := #ftK[0, #ftTot];
                                       ELSE
                                           IF #i < #ftNu AND #ftY0 + #i - #j < 48 THEN
                                               IF #ftSide[#i + 1] THEN
                                                   #ftM := #ftK[1, #ftTot] AND SHL(IN := #ftPrev[#j], N := 1);
                                               ELSE
                                                   #ftM := #ftK[2, #ftTot] AND #ftPrev[#j];
                                               END_IF;
                                           END_IF;
                                           IF #j < #ftNl AND (#CfgOrdHmi = 1 OR #i = #ftNu) THEN
                                               #ftM := #ftM OR (#ftK[3, #ftTot] AND SHR(IN := #ftCur[#j + 1], N := 1))
                                                            OR (#ftK[4, #ftTot] AND #ftCur[#j + 1]);
                                           END_IF;
                                       END_IF;
                                   END_IF;
                                   #ftCur[#j] := #ftM;
                               END_FOR;
                               FOR #j := 0 TO #ftNl DO
                                   #ftPrev[#j] := #ftCur[#j];
                               END_FOR;
                           END_FOR;
                           #ft0 := #ftCur[0];
                       END_IF;
                       IF #ftCeil <> -1 THEN
                           #bestT := 32767;
                           FOR #x := 0 TO 3 DO
                               FOR #y := 0 TO 11 DO
                                   IF #dstB = 0 THEN
                                       #id := "World".Bay0[#x, #y];
                                   ELSE
                                       #id := "World".Bay1[#x, #y];
                                   END_IF;
                                   IF #id = 0 THEN
                                       #okBal := TRUE;
                                       IF #dstB = 0 THEN
                                           #nL := "World".BalL;
                                           #nR := "World".BalR;
                                           #nF := "World".BalF;
                                           #nA := "World".BalA;
                                           IF #x <= 1 THEN #nL := #nL + 1; ELSE #nR := #nR + 1; END_IF;
                                           IF #y <= 5 THEN #nF := #nF + 1; ELSE #nA := #nA + 1; END_IF;
                                           #okBal := ABS(#nL - #nR) <= "World".CfgBalLimit
                                                     OR ABS(#nL - #nR) <= ABS("World".BalL - "World".BalR)
                                                     OR (ABS("World".BalL - "World".BalR) > "World".CfgBalLimit
                                                         AND ABS(#nL - #nR) <= "World".BalCeil);
                                           IF "World".CfgBalMode = 1 AND NOT (ABS(#nF - #nA) <= "World".CfgBalLimit
                                               OR ABS(#nF - #nA) <= ABS("World".BalF - "World".BalA))
                                           THEN
                                               #okBal := FALSE;
                                           END_IF;
                                           // v1.6: side must keep the list order feasible (tries 1 / 2)
                                           IF #okBal AND #ftCeil >= 0 AND #nL >= 0 AND #nL <= 24 THEN
                                               #ftBit := SHL(IN := DWORD#16#1, N := INT_TO_USINT(#nL));
                                               IF (#ft0 AND #ftBit) = DWORD#16#0 THEN
                                                   #okBal := FALSE;
                                               END_IF;
                                           END_IF;
                                       END_IF;
                                       IF #okBal THEN
                                           // FB1 move time in ds: max(|dx|*6 s, |dy|*2.3 s)
                                           #candT := MAX(IN1 := ABS(#x - SINT_TO_INT("World".CraneX)) * 60,
                                                         IN2 := ABS(#y - SINT_TO_INT("World".CraneY)) * 23);
                                           IF #candT < #bestT THEN
                                               #bestT := #candT;
                                               #bestX := #x;
                                               #bestY := #y;
                                           END_IF;
                                       END_IF;
                                   END_IF;
                               END_FOR;
                           END_FOR;
                       END_IF;
                   END_IF;
               END_FOR;
               IF #bestX >= 0 THEN
                   "World".Plan["World".PlanIdx].DstX := INT_TO_SINT(#bestX);
                   "World".Plan["World".PlanIdx].DstY := INT_TO_SINT(#bestY);
                   "World".Phase := 2;            // move to the new destination, then put
                   #ReplanAfterPut := TRUE;
               ELSE
                   #AlarmLatch := #AlarmLatch OR WORD#16#0080;   // bit 7 no free slot: MANUAL needed
                   #NoCellWarn := TRUE;           // v1.5 (R2-E3): shown, but not blocking -> PAUSED, MANUAL works
                   #noCell := TRUE;
               END_IF;
           ELSIF (#faultWas AND WORD#16#0005) <> 0 AND "World".Carried <> 0 THEN
               #noCell := TRUE;                   // rejected put that cannot be re-targeted: no auto retry
           END_IF;
           // A runtime fault means the yard may differ from the plan: replan from the
           // actual state. Exception: a container is on the hook - then the plan is
           // kept and resumed from the done pointer (the planner cannot start with a load).
           IF #hadFault AND "World".Carried = 0 THEN
               "World".PlanValid := FALSE;
           END_IF;
           IF #State = 5 THEN
               "World".Permit := FALSE;
               "World".CmdReady := FALSE;
               CASE #PrevState OF
                   1:  // INIT interrupted: start it again
                       #State := 1;
                       #InitStep := 0;
                   3, 7:   // was running / planning: "nakon potvrde sustav nastavlja s radom"
                       IF #Mode = 3 OR #noCell THEN
                           #State := 4;                   // PAUSED (noCell: put the container in MANUAL)
                       ELSIF "World".PlanValid THEN
                           #State := 3;
                           #Resync := TRUE;
                           #SemiTokens := 0;
                           "World".Permit := TRUE;
                       ELSE
                           #State := 7;
                           #PlanStep := 0;
                       END_IF;
                   ELSE
                       #State := #PrevState;      // READY / PAUSED / DONE
               END_CASE;
           END_IF;
       END_IF;
   END_REGION

   REGION 6 Mode selection
       IF #bAuto THEN #PendMode := 1; END_IF;
       IF #bSemi THEN #PendMode := 2; END_IF;
       IF #bManual THEN #PendMode := 3; END_IF;
       // Applied at once (also while FB1 executes: the command in FB1 always completes),
       // except during INIT.
       IF #PendMode <> 0 AND #State <> 1 THEN
           IF #PendMode = 3 AND #Mode <> 3 AND (#State = 3 OR #State = 7) THEN
               // MANUAL while running -> PAUSED; withdraw a staged plan command
               "World".Permit := FALSE;
               "World".CmdReady := FALSE;
               #State := 4;
           END_IF;
           IF #Mode = 3 AND #PendMode <> 3 AND NOT "World".Busy THEN
               // leaving MANUAL: withdraw a staged manual command
               "World".Permit := FALSE;
               "World".CmdReady := FALSE;
           END_IF;
           IF #PendMode <> #Mode THEN
               #SemiTokens := 0;
               #PendStep := FALSE;
           END_IF;
           #Mode := #PendMode;
           #PendMode := 0;
       END_IF;
   END_REGION

   REGION 7 State machine
       // ---- OFF / ON (main switch, highest priority) ----
       IF NOT "HMI_IF".SwOn THEN
           IF #State <> 0 THEN
               #OffState := #State;
               "World".Permit := FALSE;           // first Permit, then withdraw (OB30 preempts OB1)
               "World".CmdReady := FALSE;
               #SemiTokens := 0;
               #PendStep := FALSE;
               #State := 0;
           END_IF;
       ELSIF #State = 0 THEN
           IF NOT #Initialized THEN
               #State := 1;                       // first ON after PLC start -> INIT
               #InitStep := 0;
           ELSIF #OffState = 6 THEN
               #State := 6;
           ELSE
               #State := 4;                       // ON after OFF -> PAUSED (START resumes)
           END_IF;
       END_IF;

       // ---- Buttons that change the state ----
       IF "HMI_IF".SwOn THEN
           // INITIAL STATE
           // v1.5 (judge round 2 R2-J4): ignored while RUNNING / PLANNING (STOP first), so a mis-click
           // cannot reset FB1 (M, T) in the middle of a run.
           IF #bInit AND #State <> 1 AND #State <> 3 AND #State <> 7 THEN
               #State := 1;
               #InitStep := 0;
           END_IF;

           // STOP: the command in FB1 completes, a staged one is withdrawn
           IF #bStop THEN
               #PendStep := FALSE;
           END_IF;
           IF #bStop AND (#State = 3 OR #State = 7) THEN
               "World".Permit := FALSE;
               "World".CmdReady := FALSE;
               #SemiTokens := 0;
               #State := 4;
           END_IF;

           // START (AUTO / SEMI). In SEMI, NEXT STEP in READY / PAUSED acts as START + one step
           // (the latched click is executed as soon as the state is RUNNING).
           #semiGo := #PendStep AND #Mode = 2 AND (#State = 2 OR #State = 4);
           IF (#bStart OR #semiGo) AND NOT #bStop THEN
               IF NOT #Initialized THEN
                   #AlarmLatch := #AlarmLatch OR WORD#16#2000;            // bit 13 not initialized
                   #PendStep := FALSE;
               ELSIF #Mode <> 3 AND (#State = 2 OR #State = 4 OR #State = 6) THEN
                   // With a container on the hook, START is only allowed to finish the
                   // transfer that is in progress (STOP after a lift, then START).
                   #carriedOk := "World".Carried = 0;
                   IF NOT #carriedOk AND "World".PlanValid AND "World".PlanIdx >= 1
                       AND "World".PlanIdx <= "World".PlanLen AND "World".PlanIdx <= 96
                       AND "World".Phase >= 2
                   THEN
                       #carriedOk := "World".Plan["World".PlanIdx].Id = "World".Carried;
                   END_IF;
                   IF NOT #carriedOk THEN
                       #AlarmLatch := #AlarmLatch OR WORD#16#0800;        // bit 11 crane carrying
                       "HMI_IF".AlarmId := "World".Carried;
                       "HMI_IF".AlarmX := "World".CraneX;
                       "HMI_IF".AlarmY := "World".CraneY;
                       "HMI_IF".AlarmBay := "World".CraneBay;
                   ELSIF "World".PlanValid THEN
                       IF #State <> 6 THEN                                // DONE + valid plan: nothing to do
                           #State := 3;
                           #Resync := TRUE;
                           #SemiTokens := 0;
                           "World".Permit := TRUE;
                       END_IF;
                   ELSE
                       #State := 7;                                       // plan first
                       #PlanStep := 0;
                   END_IF;
               END_IF;
           END_IF;
       END_IF;

       // ---- Blocking alarm -> ALARM ----
       // blocking bits: 1, 2, 7, 8, 10, 11, 12 and every fault detected by OB30
       #blocking := (#AlarmLatch AND WORD#16#1D86) <> 0 OR "World".Fault <> 0;
       IF #NoCellWarn AND (#AlarmLatch AND WORD#16#1D06) = 0 AND "World".Fault = 0 THEN
           #blocking := FALSE;                    // v1.5 (R2-E3): bit 7 from the ACK re-target only
       END_IF;
       IF #blocking AND #State <> 0 AND #State <> 5 AND NOT (#State = 1 AND #InitStep = 0) THEN
           #PrevState := #State;
           "World".Permit := FALSE;
           "World".CmdReady := FALSE;
           #SemiTokens := 0;
           #PendStep := FALSE;
           #State := 5;
       END_IF;

       CASE #State OF
           0:  // ---------------- OFF ----------------
               ;

           1:  // ---------------- INIT (CONTRACT 3.2) ----------------
               CASE #InitStep OF
                   0:  // stop everything, clear alarms
                       "World".Permit := FALSE;
                       "World".CmdReady := FALSE;
                       "World".Fault := 0;
                       #AlarmLatch := 0;
                       #NoCellWarn := FALSE;
                       "HMI_IF".AlarmId := 0;
                       #Initialized := FALSE;
                       "World".PlanValid := FALSE;
                       #SemiTokens := 0;
                       #PendStep := FALSE;
                       #ReplanAfterPut := FALSE;
                       #OrdFallback := FALSE;
                       #InitStep := 1;

                   1:  // wait for FB1, then stage the reset command (10)
                       IF NOT "World".Busy AND NOT "World".CmdReady THEN
                           "World".NextCmd.Cmd := 10;
                           "World".NextCmd.X := 0;
                           "World".NextCmd.Y := 0;
                           "World".NextCmd.Bay := 1;
                           "World".NextCmd.Src := 4;
                           "World".NextCmd.TrIdx := 0;
                           "World".NextCmd.Phase := 0;
                           #InitSeq := "World".DoneSeq;
                           "World".Permit := TRUE;
                           "World".CmdReady := TRUE;      // last: hands the command to OB30
                           #InitStep := 2;
                       END_IF;

                   2:  // wait until OB30 reports the reset as done
                       IF "World".DoneSeq <> #InitSeq AND NOT "World".Busy AND "World".LastDone.Cmd = 10 THEN
                           "World".Permit := FALSE;
                           #InitStep := 3;
                       END_IF;

                   3:  // copy the yard and the lists, validate (all warnings except capacity)
                       // v1.4: DB10/DB11 hold the live state (region 2a). POÄŒETNO STANJE restores the
                       // data of the last load (InitBay0/1) for a repeat run, unless there is no copy yet,
                       // DB10/DB11 were edited online while no job was in progress (ExtEdit) or differ from
                       // the last mirrored state (e.g. new start values after a download): then DB10/DB11
                       // are the new yard.
                       // v1.6 (judge round 3 R3-E1 / R3-J1): cells edited with no job in progress (NewCnt)
                       // are new yard data; edits made DURING a job (obstacles, ObstCnt) only together with
                       // new lists or when >= 8 cells were rewritten. Edits written back do not count.
                       // New lists alone keep the loaded yard (InitBay) and take the new lists. The lists
                       // are always read from DB20/DB21 below.
                       #listsNew := FALSE;
                       FOR #i := 1 TO 48 DO
                           IF "From_Bay0_to_Bay1".IDs_of_the_containers[#i] <> "World".UList[#i]
                               OR "From_Bay1_to_Bay0".Bay1_IDs_of_the_containers[#i] <> "World".LList[#i]
                           THEN
                               #listsNew := TRUE;
                           END_IF;
                       END_FOR;
                       #extE := #NewCnt > 0 OR NOT #HaveInit OR (#listsNew AND #ObstCnt > 0) OR #ObstCnt >= 8;
                       FOR #x := 0 TO 3 DO
                           FOR #y := 0 TO 11 DO
                               IF "Current_state_of_Bay0".Bay0[#x, #y] <> #Snap0[#x, #y]
                                   OR "Current_state_of_Bay1".Bay1[#x, #y] <> #Snap1[#x, #y]
                               THEN
                                   #extE := TRUE;
                               END_IF;
                           END_FOR;
                       END_FOR;
                       FOR #x := 0 TO 3 DO
                           FOR #y := 0 TO 11 DO
                               IF #extE THEN
                                   #InitBay0[#x, #y] := "Current_state_of_Bay0".Bay0[#x, #y];
                                   #InitBay1[#x, #y] := "Current_state_of_Bay1".Bay1[#x, #y];
                               ELSE
                                   "Current_state_of_Bay0".Bay0[#x, #y] := #InitBay0[#x, #y];
                                   "Current_state_of_Bay1".Bay1[#x, #y] := #InitBay1[#x, #y];
                               END_IF;
                           END_FOR;
                       END_FOR;
                       #HaveInit := TRUE;
                       #ExtEdit := FALSE;
                       #JobActive := FALSE;               // v1.6: a new job starts with this load
                       #NewCnt := 0;
                       #ObstCnt := 0;
                       FOR #i := 0 TO 95 DO
                           #EditMark[#i] := FALSE;
                           #EditNew[#i] := FALSE;
                           #EditVal[#i] := 0;
                       END_FOR;
                       "HMI_IF".AlarmUId := 0;            // list IDs missing from their bay (bits 3 / 4)
                       "HMI_IF".AlarmUCnt := 0;
                       "HMI_IF".AlarmLId := 0;
                       "HMI_IF".AlarmLCnt := 0;
                       FOR #x := 0 TO 3 DO
                           FOR #y := 0 TO 11 DO
                               "World".Bay0[#x, #y] := "Current_state_of_Bay0".Bay0[#x, #y];
                               "World".Bay1[#x, #y] := "Current_state_of_Bay1".Bay1[#x, #y];
                               #Snap0[#x, #y] := "World".Bay0[#x, #y];
                               #Snap1[#x, #y] := "World".Bay1[#x, #y];
                               #tc[#x * 12 + #y] := "World".Bay0[#x, #y];
                               #tc[48 + #x * 12 + #y] := "World".Bay1[#x, #y];
                           END_FOR;
                       END_FOR;
                       "World".Carried := 0;
                       #nL := 0;                          // v1.5 (R2-J1): imbalance of the loaded data
                       #nR := 0;
                       FOR #i := 0 TO 47 DO
                           IF #tc[#i] <> 0 THEN
                               IF #i < 24 THEN #nL := #nL + 1; ELSE #nR := #nR + 1; END_IF;
                           END_IF;
                       END_FOR;
                       #BalD0 := ABS(#nL - #nR);
                       "World".BalCeil := 0;
                       "World".CraneX := "x_position";
                       "World".CraneY := "y_position";
                       "World".CraneBay := "bay_ID";

                       // cells: invalid IDs (bit 5) and duplicates (bit 6)
                       FOR #i := 0 TO 95 DO
                           #id := #tc[#i];
                           IF #id <> 0 THEN
                               IF #id < 100 OR #id > 999 THEN
                                   #AlarmLatch := #AlarmLatch OR WORD#16#0020;
                                   "HMI_IF".AlarmId := #id;
                                   "HMI_IF".AlarmBay := INT_TO_USINT(#i / 48);
                                   "HMI_IF".AlarmX := INT_TO_SINT((#i MOD 48) / 12);
                                   "HMI_IF".AlarmY := INT_TO_SINT(#i MOD 12);
                               END_IF;
                               FOR #j := #i + 1 TO 95 DO
                                   IF #tc[#j] = #id THEN
                                       #AlarmLatch := #AlarmLatch OR WORD#16#0040;
                                       "HMI_IF".AlarmId := #id;
                                       "HMI_IF".AlarmBay := INT_TO_USINT(#j / 48);
                                       "HMI_IF".AlarmX := INT_TO_SINT((#j MOD 48) / 12);
                                       "HMI_IF".AlarmY := INT_TO_SINT(#j MOD 12);
                                   END_IF;
                               END_FOR;
                           END_IF;
                       END_FOR;

                       // lists: UList 1..48 then LList 1..48 (same order as tools/crane_model.py)
                       "World".N := 0;
                       FOR #i := 1 TO 48 DO
                           "World".UList[#i] := "From_Bay0_to_Bay1".IDs_of_the_containers[#i];
                           "World".LList[#i] := "From_Bay1_to_Bay0".Bay1_IDs_of_the_containers[#i];
                           #tl[#i] := "World".UList[#i];
                           #tl[48 + #i] := "World".LList[#i];
                           IF "World".UList[#i] <> 0 THEN "World".N := "World".N + 1; END_IF;
                           IF "World".LList[#i] <> 0 THEN "World".N := "World".N + 1; END_IF;
                       END_FOR;
                       FOR #i := 1 TO 96 DO
                           #id := #tl[#i];
                           IF #id = 0 THEN
                               #ts[#i] := 2;                                  // empty entry (silent)
                           ELSIF #id < 100 OR #id > 999 THEN
                               #ts[#i] := 2;                                  // invalid ID
                               #AlarmLatch := #AlarmLatch OR WORD#16#0020;
                               "HMI_IF".AlarmId := #id;
                           ELSE
                               #found := FALSE;                               // in an earlier ACCEPTED entry?
                               FOR #j := 1 TO #i - 1 DO                       // v1.5 (R2-E1): a rejected entry does not
                                   IF #tl[#j] = #id AND #ts[#j] = 0 THEN      // kill a valid later one with the same ID
                                       #found := TRUE;
                                   END_IF;
                               END_FOR;
                               IF #found THEN
                                   #ts[#i] := 2;                              // duplicate
                                   #AlarmLatch := #AlarmLatch OR WORD#16#0040;
                                   "HMI_IF".AlarmId := #id;
                               ELSE
                                   #found := FALSE;                           // in its source bay?
                                   FOR #x := 0 TO 3 DO
                                       FOR #y := 0 TO 11 DO
                                           IF #i <= 48 THEN
                                               IF "World".Bay0[#x, #y] = #id THEN #found := TRUE; END_IF;
                                           ELSE
                                               IF "World".Bay1[#x, #y] = #id THEN #found := TRUE; END_IF;
                                           END_IF;
                                       END_FOR;
                                   END_FOR;
                                   IF #found THEN
                                       #ts[#i] := 0;                          // pending
                                   ELSE
                                       #ts[#i] := 2;
                                       IF #i <= 48 THEN
                                           #AlarmLatch := #AlarmLatch OR WORD#16#0008;  // bit 3 unload ID not in Bay 0
                                           "HMI_IF".AlarmBay := 0;
                                           IF "HMI_IF".AlarmUCnt = 0 THEN
                                               "HMI_IF".AlarmUId := #id;              // first offending ID (alarm text field)
                                           END_IF;
                                           "HMI_IF".AlarmUCnt := "HMI_IF".AlarmUCnt + 1;
                                       ELSE
                                           #AlarmLatch := #AlarmLatch OR WORD#16#0010;  // bit 4 load ID not in Bay 1
                                           "HMI_IF".AlarmBay := 1;
                                           IF "HMI_IF".AlarmLCnt = 0 THEN
                                               "HMI_IF".AlarmLId := #id;
                                           END_IF;
                                           "HMI_IF".AlarmLCnt := "HMI_IF".AlarmLCnt + 1;
                                       END_IF;
                                       "HMI_IF".AlarmId := #id;
                                       "HMI_IF".AlarmX := -1;
                                       "HMI_IF".AlarmY := -1;
                                   END_IF;
                               END_IF;
                           END_IF;
                       END_FOR;
                       #pu := 0;
                       #pl := 0;
                       FOR #i := 1 TO 48 DO
                           "World".UState[#i] := #ts[#i];
                           "World".LState[#i] := #ts[48 + #i];
                           IF #ts[#i] = 0 THEN #pu := #pu + 1; END_IF;
                           IF #ts[48 + #i] = 0 THEN #pl := #pl + 1; END_IF;
                       END_FOR;

                       // capacity (blocking, bit 7)
                       #cnt := 0;      // occupied Bay0
                       #cnt2 := 0;     // occupied Bay1
                       FOR #i := 0 TO 47 DO
                           IF #tc[#i] <> 0 THEN #cnt := #cnt + 1; END_IF;
                           IF #tc[48 + #i] <> 0 THEN #cnt2 := #cnt2 + 1; END_IF;
                       END_FOR;
                       IF #cnt2 - #pl + #pu > 48 OR #cnt - #pu + #pl > 48 THEN
                           #AlarmLatch := #AlarmLatch OR WORD#16#0080;
                           #Initialized := FALSE;
                           #PrevState := 2;
                           #State := 5;                   // ALARM; ACK -> READY (not initialized)
                       ELSE
                           // initial imbalance is only a warning (bit 0 is raised in region 4)
                           #InitStep := 4;
                       END_IF;

                   4:  // request the plan (planner idle, crane empty)
                       IF NOT "World".Busy AND #SeenSeq = "World".DoneSeq
                           AND NOT #PlanReq AND NOT #Planner.Busy AND NOT #Planner.Done AND NOT #Planner.Error
                       THEN
                           IF NOT #OrdFallback THEN       // first try: the preferred (HMI) modes
                               "World".CfgOrderMode := #CfgOrdHmi;
                               "World".CfgBalMode := #CfgBalHmi;
                               "World".BalCeil := 0;      // v1.5: step rule first
                           END_IF;
                           #OrdFallback := FALSE;
                           "World".BaseT_ds := ROUND("time" * 10.0);
                           // v1.7: the plan continues the M count of the active model (mode 0 = spec rule = World.MSpec)
                           IF "World".CfgMMode = 0 THEN
                               "World".BaseM := UDINT_TO_DINT("World".MSpec);
                           ELSE
                               "World".BaseM := UDINT_TO_DINT("number_of_manipulations");
                           END_IF;
                           #PlanCrX := "World".CraneX;
                           #PlanCrY := "World".CraneY;
                           #PlanCrBay := "World".CraneBay;
                           #PlanFinished := FALSE;
                           #PlanReq := TRUE;
                           #InitStep := 5;
                       END_IF;

                   5:  // wait for the planner
                       IF #PlanFinished THEN
                           #PlanFinished := FALSE;
                           #Initialized := TRUE;          // yard copied: MANUAL is possible even if planning failed
                           IF #PlanOk THEN
                               #State := 2;               // READY
                           ELSIF #PlanErr = 1 AND ("World".CfgOrderMode > 0 OR "World".CfgBalMode > 0) THEN
                               // dead end under the balance rule: retry with a less strict mode
                               // (order 2 -> 1 -> 0, then balance mode 1 -> 0)
                               // v1.5 (R2-J1): a ship that was loaded out of balance first gets the relaxed
                               // rule in the same order (|L-R| <= BalD0 until balanced, end balanced)
                               // v1.6 (R3-E3): World.CfgRelaxMin = ascending ceilings CfgBalLimit+1 .. BalD0
                               IF "World".CfgOrderMode > 0 AND "World".BalCeil < #BalD0 AND #BalD0 > "World".CfgBalLimit THEN
                                   IF NOT "World".CfgRelaxMin THEN
                                       "World".BalCeil := #BalD0;
                                   ELSIF "World".BalCeil = 0 THEN
                                       "World".BalCeil := "World".CfgBalLimit + 1;
                                   ELSE
                                       "World".BalCeil := "World".BalCeil + 1;
                                   END_IF;
                               ELSIF "World".CfgOrderMode > 0 THEN
                                   "World".BalCeil := 0;
                                   "World".CfgOrderMode := "World".CfgOrderMode - 1;
                               ELSE
                                   "World".BalCeil := 0;
                                   "World".CfgBalMode := 0;
                               END_IF;
                               #OrdFallback := TRUE;
                               #InitStep := 4;
                           ELSE
                               "World".PlanValid := FALSE;
                               #AlarmLatch := #AlarmLatch OR WORD#16#0100;   // bit 8 plan infeasible
                               #PrevState := 2;
                               #State := 5;
                           END_IF;
                       END_IF;

                   ELSE
                       #InitStep := 0;
               END_CASE;

           2:  // ---------------- READY ----------------
               ;   // waits for START (region above) or MANUAL commands (region 8)

           3:  // ---------------- RUNNING ----------------
               IF NOT "World".PlanValid THEN
                   #State := 7;                   // plan invalidated -> replan
                   #PlanStep := 0;
               ELSIF "World".PlanIdx > "World".PlanLen AND NOT "World".Busy AND NOT "World".CmdReady THEN
                   #cnt := 0;
                   FOR #i := 1 TO 48 DO
                       IF "World".UState[#i] = 0 THEN #cnt := #cnt + 1; END_IF;
                       IF "World".LState[#i] = 0 THEN #cnt := #cnt + 1; END_IF;
                   END_FOR;
                   IF #cnt = 0 THEN
                       "World".Permit := FALSE;
                       #AlarmLatch := #AlarmLatch OR WORD#16#8000;   // bit 15 finished (info)
                       #State := 6;               // DONE
                   ELSE
                       "World".PlanValid := FALSE;   // entries still pending -> replan
                       #State := 7;
                       #PlanStep := 0;
                   END_IF;
               END_IF;

           4:  // ---------------- PAUSED ----------------
               ;

           5:  // ---------------- ALARM ----------------
               ;   // leaves on ACK (region 5) or INIT

           6:  // ---------------- DONE ----------------
               #PendStep := FALSE;

           7:  // ---------------- PLANNING ----------------
               CASE #PlanStep OF
                   0:  // nothing may be issued while planning
                       "World".Permit := FALSE;
                       "World".CmdReady := FALSE;
                       #PlanStep := 1;
                   1:  // wait for FB1 and an idle planner, then request
                       // NOT Busy first, then SeenSeq = DoneSeq: list states include the last PUT
                       IF NOT "World".Busy AND #SeenSeq = "World".DoneSeq AND NOT #PlanReq AND NOT #Planner.Busy
                           AND NOT #Planner.Done AND NOT #Planner.Error
                       THEN
                           IF "World".Carried <> 0 THEN
                               // the planner needs an empty hook: put it down in MANUAL first
                               #AlarmLatch := #AlarmLatch OR WORD#16#0800;   // bit 11
                               "HMI_IF".AlarmId := "World".Carried;
                               #PrevState := 4;
                               #State := 5;
                           ELSE
                               // Pending entries whose container is no longer in its source bay
                               // (MANUAL moves, online DB10/DB11 edits): done if it is in the
                               // destination bay, otherwise skipped with warning bit 3 / 4.
                               FOR #i := 1 TO 48 DO
                                   FOR #k := 1 TO 2 DO
                                       IF #k = 1 THEN
                                           #id := "World".UList[#i];
                                           #found := "World".UState[#i] = 0;
                                       ELSE
                                           #id := "World".LList[#i];
                                           #found := "World".LState[#i] = 0;
                                       END_IF;
                                       IF #found THEN
                                           #found0 := FALSE;
                                           #found1 := FALSE;
                                           FOR #x := 0 TO 3 DO
                                               FOR #y := 0 TO 11 DO
                                                   IF "World".Bay0[#x, #y] = #id THEN #found0 := TRUE; END_IF;
                                                   IF "World".Bay1[#x, #y] = #id THEN #found1 := TRUE; END_IF;
                                               END_FOR;
                                           END_FOR;
                                           IF #k = 1 AND NOT #found0 THEN
                                               IF #found1 THEN
                                                   "World".UState[#i] := 1;
                                               ELSE
                                                   "World".UState[#i] := 2;
                                                   #AlarmLatch := #AlarmLatch OR WORD#16#0008;
                                                   "HMI_IF".AlarmId := #id;
                                                   "HMI_IF".AlarmBay := 0;
                                                   "HMI_IF".AlarmX := -1;
                                                   "HMI_IF".AlarmY := -1;
                                               END_IF;
                                           ELSIF #k = 2 AND NOT #found1 THEN
                                               IF #found0 THEN
                                                   "World".LState[#i] := 1;
                                               ELSE
                                                   "World".LState[#i] := 2;
                                                   #AlarmLatch := #AlarmLatch OR WORD#16#0010;
                                                   "HMI_IF".AlarmId := #id;
                                                   "HMI_IF".AlarmBay := 1;
                                                   "HMI_IF".AlarmX := -1;
                                                   "HMI_IF".AlarmY := -1;
                                               END_IF;
                                           END_IF;
                                       END_IF;
                                   END_FOR;
                               END_FOR;
                               IF NOT #OrdFallback THEN   // first try: the preferred (HMI) modes
                                   "World".CfgOrderMode := #CfgOrdHmi;
                                   "World".CfgBalMode := #CfgBalHmi;
                                   "World".BalCeil := 0;  // v1.5: step rule first
                               END_IF;
                               #OrdFallback := FALSE;
                               "World".BaseT_ds := ROUND("time" * 10.0);
                               // v1.7: the plan continues the M count of the active model (mode 0 = spec rule = World.MSpec)
                               IF "World".CfgMMode = 0 THEN
                                   "World".BaseM := UDINT_TO_DINT("World".MSpec);
                               ELSE
                                   "World".BaseM := UDINT_TO_DINT("number_of_manipulations");
                               END_IF;
                               #PlanCrX := "World".CraneX;
                               #PlanCrY := "World".CraneY;
                               #PlanCrBay := "World".CraneBay;
                               #PlanFinished := FALSE;
                               #PlanReq := TRUE;
                               #PlanStep := 2;
                           END_IF;
                       END_IF;
                   2:  // wait for the result
                       IF #PlanFinished THEN
                           #PlanFinished := FALSE;
                           IF #PlanOk THEN
                               IF #Mode = 3 THEN
                                   #State := 4;
                               ELSE
                                   #State := 3;
                                   #Resync := TRUE;
                                   #SemiTokens := 0;
                                   "World".Permit := TRUE;
                               END_IF;
                           ELSIF #PlanErr = 1 AND ("World".CfgOrderMode > 0 OR "World".CfgBalMode > 0) THEN
                               // dead end: retry with a less strict mode (see INIT step 5)
                               // v1.5 (R2-J1): a ship that was loaded out of balance first gets the relaxed
                               // rule in the same order (|L-R| <= BalD0 until balanced, end balanced)
                               // v1.6 (R3-E3): World.CfgRelaxMin = ascending ceilings CfgBalLimit+1 .. BalD0
                               IF "World".CfgOrderMode > 0 AND "World".BalCeil < #BalD0 AND #BalD0 > "World".CfgBalLimit THEN
                                   IF NOT "World".CfgRelaxMin THEN
                                       "World".BalCeil := #BalD0;
                                   ELSIF "World".BalCeil = 0 THEN
                                       "World".BalCeil := "World".CfgBalLimit + 1;
                                   ELSE
                                       "World".BalCeil := "World".BalCeil + 1;
                                   END_IF;
                               ELSIF "World".CfgOrderMode > 0 THEN
                                   "World".BalCeil := 0;
                                   "World".CfgOrderMode := "World".CfgOrderMode - 1;
                               ELSE
                                   "World".BalCeil := 0;
                                   "World".CfgBalMode := 0;
                               END_IF;
                               #OrdFallback := TRUE;
                               #PlanStep := 1;
                           ELSE
                               "World".PlanValid := FALSE;
                               #AlarmLatch := #AlarmLatch OR WORD#16#0100;   // bit 8 plan infeasible
                               #PrevState := 4;
                               #State := 5;
                           END_IF;
                       END_IF;
                   ELSE
                       #PlanStep := 0;
               END_CASE;

           ELSE
               #State := 0;
       END_CASE;
   END_REGION

   REGION 8 New plan: done pointer, staging cursor, skip rule
       // Runs once when a plan was just accepted (INIT step 5 / PLANNING step 2 set PlanFinished := FALSE
       // and PlanOk = TRUE in this cycle). The pointers are set from the plan-time crane position.
       IF #PlanOk AND NOT #PlanFinished AND NOT #PlanReq AND "World".PlanValid
           AND ((#State = 2 AND #InitStep = 5) OR ((#State = 3 OR #State = 4) AND #PlanStep = 2))
       THEN
           IF "World".PlanLen > 96 THEN
               "World".PlanLen := 96;
           END_IF;
           // Skip rule (CONTRACT 3.4): move-to-src is skipped when the crane is already there
           FOR #i := 1 TO "World".PlanLen DO
               IF #i = 1 THEN
                   #found := #PlanCrX = "World".Plan[1].SrcX AND #PlanCrY = "World".Plan[1].SrcY
                             AND #PlanCrBay = "World".Plan[1].SrcBay;
               ELSE
                   #found := "World".Plan[#i - 1].DstX = "World".Plan[#i].SrcX
                             AND "World".Plan[#i - 1].DstY = "World".Plan[#i].SrcY
                             AND "World".Plan[#i - 1].DstBay = "World".Plan[#i].SrcBay;
               END_IF;
               IF #found THEN
                   #FirstPh[#i] := 1;
               ELSE
                   #FirstPh[#i] := 0;
               END_IF;
           END_FOR;
           "World".PlanIdx := 1;
           IF "World".PlanLen >= 1 THEN
               "World".Phase := #FirstPh[1];
           ELSE
               "World".Phase := 0;
           END_IF;
           "World".StageIdx := 1;
           "World".StagePhase := "World".Phase;
           #ReplanAfterPut := FALSE;
           #InitStep := 6;                        // INIT finished
           #PlanStep := 3;                        // PLANNING finished
           #PlanOk := FALSE;                      // consumed
       END_IF;
   END_REGION

   REGION 9 Staging: AUTO / SEMI plan commands, MANUAL commands
       // ---- AUTO / SEMI: next plan command (at most one staged ahead of FB1) ----
       IF #State = 3 AND #Mode <> 3 AND "World".PlanValid AND "World".Permit THEN
           // After START / ACK: continue exactly from the done pointer
           // (NOT Busy first, then SeenSeq = DoneSeq: every completion is already counted)
           IF #Resync AND NOT "World".Busy AND #SeenSeq = "World".DoneSeq AND NOT "World".CmdReady THEN
               "World".StageIdx := "World".PlanIdx;
               "World".StagePhase := "World".Phase;
               #Resync := FALSE;
           END_IF;

           // SEMI: one click = one command (or the rest of one transfer); the click is latched
           // (PendStep) and executed as soon as FB1 has finished the previous command
           IF #Mode = 2 AND #PendStep AND NOT #Resync AND #SemiTokens = 0
               AND NOT "World".Busy AND NOT "World".CmdReady
           THEN
               #PendStep := FALSE;
               IF "HMI_IF".CfgSemiPerTransfer THEN
                   #SemiTokens := 4 - USINT_TO_INT("World".StagePhase);
               ELSE
                   #SemiTokens := 1;
               END_IF;
           END_IF;

           IF NOT #Resync AND NOT "World".CmdReady
               AND "World".StageIdx >= 1 AND "World".StageIdx <= "World".PlanLen AND "World".StageIdx <= 96
               AND (#Mode = 1 OR #SemiTokens > 0)
           THEN
               #tr := "World".Plan["World".StageIdx];
               CASE "World".StagePhase OF
                   0:  "World".NextCmd.Cmd := 3;          // move to source
                   1:  "World".NextCmd.Cmd := 1;          // lift
                   2:  "World".NextCmd.Cmd := 3;          // move to destination
                   ELSE
                       "World".NextCmd.Cmd := 2;          // put down
               END_CASE;
               IF "World".StagePhase <= 1 THEN
                   "World".NextCmd.X := #tr.SrcX;
                   "World".NextCmd.Y := #tr.SrcY;
                   "World".NextCmd.Bay := #tr.SrcBay;
               ELSE
                   "World".NextCmd.X := #tr.DstX;
                   "World".NextCmd.Y := #tr.DstY;
                   "World".NextCmd.Bay := #tr.DstBay;
               END_IF;
               "World".NextCmd.Src := #Mode;              // 1 AUTO, 2 SEMI
               "World".NextCmd.TrIdx := "World".StageIdx;
               "World".NextCmd.Phase := "World".StagePhase;
               "World".CmdReady := TRUE;                  // last: hands the command to OB30

               // advance the staging cursor
               IF "World".StagePhase >= 3 THEN
                   "World".StageIdx := "World".StageIdx + 1;
                   IF "World".StageIdx <= "World".PlanLen AND "World".StageIdx <= 96 THEN
                       "World".StagePhase := #FirstPh["World".StageIdx];
                   ELSE
                       "World".StagePhase := 0;
                   END_IF;
               ELSE
                   "World".StagePhase := "World".StagePhase + 1;
               END_IF;
               IF #Mode = 2 AND #SemiTokens > 0 THEN
                   #SemiTokens := #SemiTokens - 1;
               END_IF;
           END_IF;
       END_IF;

       // ---- MANUAL: command from the HMI fields ----
       IF #bManExec AND #Mode = 3 AND "HMI_IF".SwOn THEN
           IF NOT #Initialized THEN
               #AlarmLatch := #AlarmLatch OR WORD#16#2000;            // bit 13 not initialized
           ELSIF (#State = 2 OR #State = 4 OR #State = 6) AND NOT #blocking
               AND NOT "World".Busy AND NOT "World".CmdReady
           THEN
               IF NOT ("HMI_IF".ManCmd = 1 OR "HMI_IF".ManCmd = 2 OR "HMI_IF".ManCmd = 3 OR "HMI_IF".ManCmd = 10)
                   OR ("HMI_IF".ManCmd = 3 AND ("HMI_IF".ManX < 0 OR "HMI_IF".ManX > 3
                       OR "HMI_IF".ManY < 0 OR "HMI_IF".ManY > 11 OR "HMI_IF".ManBay > 1))
               THEN
                   // invalid manual input: warning, the command is dropped
                   #AlarmLatch := #AlarmLatch OR WORD#16#0200;        // bit 9
                   "HMI_IF".AlarmId := 0;
                   "HMI_IF".AlarmX := "HMI_IF".ManX;
                   "HMI_IF".AlarmY := "HMI_IF".ManY;
                   "HMI_IF".AlarmBay := "HMI_IF".ManBay;
               ELSIF "HMI_IF".ManCmd = 3 AND "HMI_IF".ManX = "World".CraneX AND "HMI_IF".ManY = "World".CraneY
                   AND "HMI_IF".ManBay = "World".CraneBay
               THEN
                   ;   // zero-distance move: FB1 would add 1 manipulation for nothing -> dropped
               ELSE
                   "World".NextCmd.Cmd := "HMI_IF".ManCmd;
                   IF "HMI_IF".ManCmd = 3 THEN
                       "World".NextCmd.X := "HMI_IF".ManX;
                       "World".NextCmd.Y := "HMI_IF".ManY;
                       "World".NextCmd.Bay := "HMI_IF".ManBay;
                   ELSIF "HMI_IF".ManCmd = 10 THEN
                       "World".NextCmd.X := 0;
                       "World".NextCmd.Y := 0;
                       "World".NextCmd.Bay := 1;
                   ELSE    // lift / put: where the crane is
                       "World".NextCmd.X := "World".CraneX;
                       "World".NextCmd.Y := "World".CraneY;
                       "World".NextCmd.Bay := "World".CraneBay;
                   END_IF;
                   "World".NextCmd.Src := 3;
                   "World".NextCmd.TrIdx := 0;
                   "World".NextCmd.Phase := 0;
                   "World".Permit := TRUE;
                   "World".CmdReady := TRUE;              // last
               END_IF;
           END_IF;
       END_IF;
   END_REGION

   REGION 10 Discard a planner result nobody waits for (STOP / OFF / INIT during planning)
       IF #PlanFinished AND NOT (#State = 1 AND #InitStep = 5) AND NOT (#State = 7 AND #PlanStep = 2) THEN
           #PlanFinished := FALSE;
           #PlanOk := FALSE;
           "World".PlanValid := FALSE;
       END_IF;
   END_REGION

   REGION 11 Alarm history (ring, [0] newest)
       #newBits := #AlarmLatch AND NOT #AlarmPrev;
       IF #newBits <> 0 THEN
           FOR #b := 0 TO 15 DO
               IF (#newBits AND SHL(IN := WORD#16#0001, N := INT_TO_UINT(#b))) <> 0 THEN
                   FOR #k := 15 TO 1 BY -1 DO
                       "HMI_IF".AlarmHist[#k] := "HMI_IF".AlarmHist[#k - 1];
                       #AlarmHistM[#k] := #AlarmHistM[#k - 1];
                       #AlarmHistT[#k] := #AlarmHistT[#k - 1];
                   END_FOR;
                   "HMI_IF".AlarmHist[0] := #b;
                   #AlarmHistM[0] := "World".MSpec;   // v1.7: spec-rule M (primary)
                   #AlarmHistT[0] := "time";
                   "HMI_IF".AlarmHistSeq := "HMI_IF".AlarmHistSeq + 1;
               END_IF;
           END_FOR;
       END_IF;
       #AlarmPrev := #AlarmLatch;
   END_REGION

   REGION 12 HMI indicators (every cycle)
       // ---- state, mode, lamps ----
       #blocking := (#AlarmLatch AND WORD#16#1D86) <> 0 OR "World".Fault <> 0;
       IF #NoCellWarn AND (#AlarmLatch AND WORD#16#1D06) = 0 AND "World".Fault = 0 THEN
           #blocking := FALSE;                    // v1.5 (R2-E3): bit 7 from the ACK re-target only
       END_IF;
       "HMI_IF".State := #State;
       "HMI_IF".Mode := #Mode;
       "HMI_IF".LampOn := "HMI_IF".SwOn;
       "HMI_IF".LampOff := NOT "HMI_IF".SwOn;
       "HMI_IF".LampReady := "HMI_IF".SwOn AND #Initialized AND NOT #blocking
                             AND (#State = 2 OR #State = 3 OR #State = 4 OR #State = 6);
       "HMI_IF".LampAuto := #Mode = 1;
       "HMI_IF".LampSemi := #Mode = 2;
       "HMI_IF".LampManual := #Mode = 3;
       "HMI_IF".LampRunning := #State = 3;
       "HMI_IF".LampAlarm := (#AlarmLatch AND WORD#16#7FFF) <> 0;
       "HMI_IF".LampDone := #State = 6;
       "HMI_IF".Initialized := #Initialized;
       "HMI_IF".CraneBusy := "World".Busy;
       "HMI_IF".Planning := #State = 7 OR #Planner.Busy;
       "HMI_IF".StepWaiting := #State = 3 AND #Mode = 2 AND #SemiTokens = 0
                               AND NOT "World".Busy AND NOT "World".CmdReady
                               AND "World".StageIdx <= "World".PlanLen;
       "HMI_IF".AlarmWord := #AlarmLatch;
       "HMI_IF".AlarmAckWord := NOT #AlarmLatch;  // WinCC PLC acknowledgement: cleared bit = acknowledged
       "HMI_IF".OrderModeAct := "World".CfgOrderMode;
       // v1.4: the plan does not follow the preferred (HMI) order / balance mode because that mode is
       // provably infeasible (FB11 exact check) -> warning AlarmWord2 bit 0 (HMI alarm, no stop)
       "HMI_IF".OrderFallback := #Initialized AND "World".PlanValid
                                 AND ("World".CfgOrderMode <> #CfgOrdHmi OR "World".CfgBalMode <> #CfgBalHmi);
       IF "HMI_IF".OrderFallback THEN
           "HMI_IF".AlarmWord2 := WORD#16#0001;
       ELSE
           "HMI_IF".AlarmWord2 := WORD#16#0000;
       END_IF;
       // v1.5 (R2-J1): the plan uses the relaxed balance rule (ship loaded out of balance) -> bit 1
       IF #Initialized AND "World".PlanValid AND "World".BalCeil > "World".CfgBalLimit THEN
           "HMI_IF".AlarmWord2 := "HMI_IF".AlarmWord2 OR WORD#16#0002;
       END_IF;
       "HMI_IF".OB30Ticks := "World".OB30Ticks;

       // ---- score: M, T and J = 0.5*T/(76*N) + 0.5*M/(4*N) ----
       // v1.7: primary M / J = spec rule (diagonal x+y move = 2 M), counted by OB30 in World.MSpec.
       // FB1's own counter MD107 (+1 per move command) stays visible as MFb1 / JFb1 (secondary).
       "HMI_IF".M := "World".MSpec;
       "HMI_IF".MFb1 := "number_of_manipulations";
       "HMI_IF".T := "time";
       "HMI_IF".N := "World".N;
       IF "World".N > 0 THEN
           #rN := INT_TO_REAL("World".N);
           "HMI_IF".J := 0.5 * "time" / (76.0 * #rN) + 0.5 * UDINT_TO_REAL("World".MSpec) / (4.0 * #rN);
           "HMI_IF".JFb1 := 0.5 * "time" / (76.0 * #rN) + 0.5 * UDINT_TO_REAL("number_of_manipulations") / (4.0 * #rN);
       ELSE
           "HMI_IF".J := 0.0;
           "HMI_IF".JFb1 := 0.0;
       END_IF;
       "HMI_IF".MSpec := "HMI_IF".M;           // compatibility copies (= primary spec values)
       "HMI_IF".JSpec := "HMI_IF".J;
       "HMI_IF".PredM := "World".PredM;
       "HMI_IF".PredT := DINT_TO_REAL("World".PredT_ds) / 10.0;
       "HMI_IF".PredJ := "World".PredJ;
       "HMI_IF".PlanVariant := "World".PlanVariant;
       // v1.3: greedy J, lower bound, gap to the bound, improve-phase progress
       "HMI_IF".PredJ0 := "World".PredJ0;
       "HMI_IF".LbJ := "World".LbJ;
       IF "World".LbJ > 0.0 THEN
           "HMI_IF".GapPct := ("World".PredJ / "World".LbJ - 1.0) * 100.0;
       ELSE
           "HMI_IF".GapPct := 0.0;
       END_IF;
       IF "World".PredJ0 > 0.0 THEN
           "HMI_IF".ImpGainPct := (1.0 - "World".PredJ / "World".PredJ0) * 100.0;
       ELSE
           "HMI_IF".ImpGainPct := 0.0;
       END_IF;
       "HMI_IF".ImpEvals := "World".ImpEvals;
       "HMI_IF".SlotAccepts := "World".SlotAccepts;
       IF #Planner.Busy AND #Planner.ImpActive AND "World".CfgImproveEvals > 0 THEN
           "HMI_IF".PlanProgress := DINT_TO_INT(#Planner.ImpEvals * 100 / "World".CfgImproveEvals);
       ELSIF #Planner.Busy THEN
           "HMI_IF".PlanProgress := 0;
       ELSE
           "HMI_IF".PlanProgress := 100;
       END_IF;

       // ---- crane ----
       "HMI_IF".CraneX := "World".CraneX;
       "HMI_IF".CraneY := "World".CraneY;
       "HMI_IF".CraneBay := "World".CraneBay;
       IF "World".CraneBay = 0 THEN
           "HMI_IF".CraneGX := SINT_TO_INT("World".CraneX) + 6;
       ELSE
           "HMI_IF".CraneGX := SINT_TO_INT("World".CraneX);
       END_IF;
       "HMI_IF".Carried := "World".Carried;

       // ---- current command and transfer ----
       IF "World".Busy THEN
           #cur := "World".ActCmd;
       ELSIF "World".CmdReady THEN
           #cur := "World".NextCmd;
       ELSE
           #cur := "World".LastDone;
       END_IF;
       "HMI_IF".CurCmd := #cur.Cmd;
       "HMI_IF".CurX := #cur.X;
       "HMI_IF".CurY := #cur.Y;
       "HMI_IF".CurBay := #cur.Bay;
       "HMI_IF".CurPhase := "World".Phase;
       #curValid := "World".PlanValid AND "World".PlanIdx >= 1 AND "World".PlanIdx <= "World".PlanLen
                    AND "World".PlanIdx <= 96 AND (#State = 3 OR #State = 4 OR #State = 5);
       IF #curValid THEN
           #tr := "World".Plan["World".PlanIdx];
           "HMI_IF".CurId := #tr.Id;
           "HMI_IF".CurKind := #tr.Kind;
       ELSE
           "HMI_IF".CurId := "World".Carried;
           "HMI_IF".CurKind := 0;
       END_IF;

